// TIA Portal project "Lab_4" (V16)

(* hardware
DEVICE "S7300/ET200M station_1"  S7-300 station
   slot 0: "Rail_0"  Rail  6ES7 390-1***0-0AA0
   slot 2: "PLC_1"  CPU 315-2 DP  6ES7 315-2AG10-0AB0  V2.6
      slot 0: "MPI interface_1"  X1
      slot 1: "DP interface_1"  X2
*)

// ===== PLC "PLC_1"  CPU 315-2 DP =====

VAR_GLOBAL   // PLC tag table "Default tag table"
   "Tag_1" AT %MB20 : Byte;
   "Tag_2" AT %M20.7 : Bool;
   "Tag_3" AT %M20.0 : Bool;
   "Tag_4" AT %MD12 : DWord;
   "Tag_5" AT %M20.1 : Bool;
   "Tag_6" AT %M20.2 : Bool;
   "Tag_7" AT %MW10 : Word;
   "Tag_8" AT %MW4 : Word;
   "Tag_9" AT %MW30 : Word;
   "Tag_10" AT %MD32 : Real;
   "Tag_11" AT %MD36 : Real;
   "Tag_12" AT %MB40 : Byte;
   "Tag_13" AT %MD44 : Real;
END_VAR

FUNCTION "FC6" : Void   // FC6, STL
{ S7_Optimized_Access := 'FALSE' }
VERSION : 0.1
   VAR_INPUT
      ACQ : Word;
      SS : Real;
      SI : Real;
      "a" : Real;
      "b" : Real;
   END_VAR
   VAR_OUTPUT
      STAT : Byte;
      VAL : Real;
   END_VAR
BEGIN

REGION Network 1
         L     0;  // Initializations
         T     "Tag_1";
         T     #STAT;
         L     #ACQ;  // Load acquired value
         T     "Tag_7";  // Save in MW10
         L     W#16#7FFF;  // If acquisition error
         ==I;
         JC    ESCI;  // Return
         L     "Tag_7";  // Load acquired value
         ITD;  // Convert to 32-bit
         DTR;  // Convert to real
         L     #"a";  // Load parameter a
         *R;  // Multiply
         L     #"b";  // Load parameter b
         +R;  // Sum
         T     #VAL;  // Copy converted value on output parameter VAL
         T     "Tag_4";  // Save converted value in MD12
         L     #SS;  // Load high threshold
         >R;  // Comparison
         =     "Tag_5";  // Copy result of comparison in M20.1
         L     #SI;  // Load low threashold
         L     "Tag_4";  // Load converted value
         >R;  // Comparison
         =     "Tag_6";  // Copy result of comparison in M20.2
         L     "Tag_1";
         L     0;
         <>I;  // Check if MB20 not 0
         =     "Tag_2";  // Report in cumulative error bit
         L     "Tag_1";  // Load status byte
         T     #STAT;  // Copy on output parameter STAT
         BEU;
   ESCI: L     DW#16#FFFFFFFF;  // Load error constant
         T     #VAL;  // Copy on parameter VAL
         SET;  // Put RLO =1
         =     "Tag_3";  // Copy to M20.0 and M20.7
         =     "Tag_2";
         L     "Tag_1";  // Load status byte
         T     #STAT;  // Copy on output parameter STAT
END_REGION
END_FUNCTION

ORGANIZATION_BLOCK "Main"   // OB1, STL
TITLE = "Main Program Sweep (Cycle)"
{ S7_Optimized_Access := 'FALSE' }
VERSION : 0.1
   VAR_TEMP
      OB1_EV_CLASS : Byte;   // Bits 0-3 = 1 (Coming event), Bits 4-7 = 1 (Event class 1)
      OB1_SCAN_1 : Byte;   // 1 (Cold restart scan 1 of OB 1), 3 (Scan 2-n of OB 1)
      OB1_PRIORITY : Byte;   // Priority of OB Execution
      OB1_OB_NUMBR : Byte;   // 1 (Organization block 1, OB1)
      OB1_RESERVED_1 : Byte;   // Reserved for system
      OB1_RESERVED_2 : Byte;   // Reserved for system
      OB1_PREV_CYCLE : Int;   // Cycle time of previous OB1 scan (milliseconds)
      OB1_MIN_CYCLE : Int;   // Minimum cycle time of OB1 (milliseconds)
      OB1_MAX_CYCLE : Int;   // Maximum cycle time of OB1 (milliseconds)
      OB1_DATE_TIME : Date_And_Time;   // Date and time OB1 started
   END_VAR
BEGIN

REGION Network 1
         CALL  "FC6"
         ( ACQ  := "Tag_9",
           SS   := "Tag_10",
           SI   := "Tag_11",
           "a"  := 2.0,
           "b"  := 5.0,
           STAT := "Tag_12",
           VAL  := "Tag_13"
         );
END_REGION
END_ORGANIZATION_BLOCK